FUNCTION F_CheckHighNibbleLEDState : BOOL
VAR_IN_OUT CONSTANT
    nValue: BYTE;
END_VAR
VAR_INPUT
    bFlashOn: BOOL;
END_VAR
VAR
    nNibble: BYTE;
END_VAR

nNibble := SHR(nValue, 4);
F_CheckHighNibbleLEDState := (nNibble <> BYTE#0) AND ((nNibble <> BYTE#3) OR bFlashOn);

END_FUNCTION

(* stored: Version 1.1.0.1
   POU F_CheckHighNibbleLEDState: Id {4b91c791-0e9f-036d-15df-1e0a57ceba05}, SpecialFunc None *)
